Fanuc KAREL source: KA00059.KL

PROGRAM KA00059
%NOLOCKGROUP
VAR
  SRC: POSITION
  DST: ARRAY[2] OF BYTE
BEGIN
  DST[1] = SRC
END KA00059
